(* IEC 61131-3 sources: tgbot_base/CodeSys, 8 files *)

(* ---- GVL_IO.st ---- *)
VAR_GLOBAL
	(* ===================== MODE AND COMMON ===================== *)
	I_ModeManual AT %IX0.0 : BOOL; (* Manual/Automatic selector switch: 1 = Manual, 0 = Automatic *)
	HMI_Auto_Start : BOOL; (* HMI request to enable automatic sequence when in automatic mode *)
	HMI_ResetFaults : BOOL; (* HMI command to reset latched emergency conditions *)

	(* ===================== HMI MANUAL COMMANDS ===================== *)
	HMI_Fan1_Start : BOOL; (* Manual start for Local Fan 1 *)
	HMI_Fan2_Start : BOOL; (* Manual start for Local Fan 2 *)
	HMI_Fan3_Start : BOOL; (* Manual start for Local Fan 3 *)
	HMI_Fan4_Start : BOOL; (* Manual start for Local Fan 4 *)
	HMI_Fan5_Start : BOOL; (* Manual start for Local Fan 5 *)
	HMI_TransportFan_Start : BOOL; (* Manual start for Transport Fan *)
	HMI_Screw_Start : BOOL; (* Manual start for Screw Conveyor *)
	HMI_Vibrator1_Start : BOOL; (* Manual start for Vibrator 1 *)
	HMI_Vibrator2_Start : BOOL; (* Manual start for Vibrator 2 *)
	HMI_Hydraulic_Open : BOOL; (* Manual open command for Hydraulic Hatch *)
	HMI_Hydraulic_Close : BOOL; (* Manual close command for Hydraulic Hatch *)

	(* ===================== PHYSICAL INPUTS (FAULTS, LIMITS) ===================== *)
	(* VFD Faults for Local Fans *)
	I_Fan1_VFD_Fault AT %IX1.0 : BOOL; (* VFD fault for Local Fan 1 *)
	I_Fan2_VFD_Fault AT %IX1.1 : BOOL; (* VFD fault for Local Fan 2 *)
	I_Fan3_VFD_Fault AT %IX1.2 : BOOL; (* VFD fault for Local Fan 3 *)
	I_Fan4_VFD_Fault AT %IX1.3 : BOOL; (* VFD fault for Local Fan 4 *)
	I_Fan5_VFD_Fault AT %IX1.4 : BOOL; (* VFD fault for Local Fan 5 *)

	(* VFD Faults for other mechanisms — keep within byte 1 for example mapping *)
	I_TransportFan_VFD_Fault AT %IX1.5 : BOOL; (* VFD fault for Transport Fan *)
	I_Screw_VFD_Fault AT %IX1.6 : BOOL; (* VFD fault for Screw Conveyor *)
	I_Vibrator1_VFD_Fault AT %IX1.7 : BOOL; (* VFD fault for Vibrator 1 (if applicable) *)
	I_Vibrator2_VFD_Fault AT %IX3.0 : BOOL; (* VFD fault for Vibrator 2 (if applicable); mapped to input byte 3 bit 0 *)

	(* Circuit breaker trips (as per requirement: only vibrators and hydraulic motor) *)
	I_Vibrator1_CB_Trip AT %IX2.0 : BOOL; (* Circuit breaker trip for Vibrator 1 *)
	I_Vibrator2_CB_Trip AT %IX2.1 : BOOL; (* Circuit breaker trip for Vibrator 2 *)
	I_Hydraulic_CB_Trip AT %IX2.2 : BOOL; (* Circuit breaker trip for Hydraulic Power Unit/Motor *)

	(* Hydraulic hatch limit switches *)
	I_Hatch_Open_LS AT %IX2.3 : BOOL; (* Hydraulic Hatch OPEN position limit switch *)
	I_Hatch_Closed_LS AT %IX2.4 : BOOL; (* Hydraulic Hatch CLOSED position limit switch *)

	(* ===================== PHYSICAL OUTPUTS (COMMANDS) ===================== *)
	Q_Fan1_Run AT %QX0.0 : BOOL; (* Run command for Local Fan 1 *)
	Q_Fan2_Run AT %QX0.1 : BOOL; (* Run command for Local Fan 2 *)
	Q_Fan3_Run AT %QX0.2 : BOOL; (* Run command for Local Fan 3 *)
	Q_Fan4_Run AT %QX0.3 : BOOL; (* Run command for Local Fan 4 *)
	Q_Fan5_Run AT %QX0.4 : BOOL; (* Run command for Local Fan 5 *)
	Q_TransportFan_Run AT %QX0.5 : BOOL; (* Run command for Transport Fan *)
	Q_Screw_Run AT %QX0.6 : BOOL; (* Run command for Screw Conveyor *)
	Q_Vibrator1_Run AT %QX1.0 : BOOL; (* Run command for Vibrator 1 *)
	Q_Vibrator2_Run AT %QX1.1 : BOOL; (* Run command for Vibrator 2 *)
	Q_Hydraulic_Open AT %QX1.2 : BOOL; (* Open command for Hydraulic Hatch actuator *)
	Q_Hydraulic_Close AT %QX1.3 : BOOL; (* Close command for Hydraulic Hatch actuator *)

	(* ===================== STATUS / DIAGNOSTICS FOR HMI ===================== *)
	Status_ModeManual : BOOL; (* Current mode: TRUE = Manual, FALSE = Automatic *)
	Status_AutoEnabled : BOOL; (* Auto sequence enable status *)
	Status_EmergencyActive : BOOL; (* Emergency latch active *)

	Status_Fan1_Running : BOOL; (* Status of Local Fan 1 command *)
	Status_Fan2_Running : BOOL; (* Status of Local Fan 2 command *)
	Status_Fan3_Running : BOOL; (* Status of Local Fan 3 command *)
	Status_Fan4_Running : BOOL; (* Status of Local Fan 4 command *)
	Status_Fan5_Running : BOOL; (* Status of Local Fan 5 command *)
	Status_TransportFan_Running : BOOL; (* Status of Transport Fan command *)
	Status_Screw_Running : BOOL; (* Status of Screw Conveyor command *)
	Status_Vibrator1_Running : BOOL; (* Status of Vibrator 1 command *)
	Status_Vibrator2_Running : BOOL; (* Status of Vibrator 2 command *)
	Status_Hydraulic_Busy : BOOL; (* Hydraulic Hatch actuator active (open or close) *)
END_VAR

(* ---- FB_AutoControl.st ---- *)
FUNCTION_BLOCK FB_AutoControl
VAR_INPUT
	AutoMode : BOOL; (* TRUE when selector is in automatic mode *)
	AutoStartRequest : BOOL; (* HMI request to enable automatic sequence *)
	GlobalPermit : BOOL; (* Permit from emergency handling; must be TRUE to run *)
END_VAR
VAR_OUTPUT
	AutoEnabled : BOOL; (* Auto mode active and permitted *)
	Fan1Start : BOOL; (* Auto start command for Local Fan 1 *)
	Fan2Start : BOOL; (* Auto start command for Local Fan 2 *)
	Fan3Start : BOOL; (* Auto start command for Local Fan 3 *)
	Fan4Start : BOOL; (* Auto start command for Local Fan 4 *)
	Fan5Start : BOOL; (* Auto start command for Local Fan 5 *)
	TransportFanStart : BOOL; (* Auto start command for Transport Fan *)
	ScrewStart : BOOL; (* Auto start command for Screw Conveyor *)
	Vibrator1Start : BOOL; (* Auto start command for Vibrator 1 *)
	Vibrator2Start : BOOL; (* Auto start command for Vibrator 2 *)
END_VAR
VAR
	tFan2 : TON;
	tFan3 : TON;
	tFan4 : TON;
	tFan5 : TON;
	tTransport : TON;
	tScrew : TON;
	tVibrators : TON;
	sequenceEnabled : BOOL;
END_VAR

(* Determine if automatic control is enabled *)
sequenceEnabled := AutoMode AND AutoStartRequest AND GlobalPermit;
AutoEnabled := sequenceEnabled;

(* Progressive start delays for fans 2..5 from AutoEnabled *)
tFan2(IN := sequenceEnabled, PT := T#1S);
tFan3(IN := sequenceEnabled, PT := T#2S);
tFan4(IN := sequenceEnabled, PT := T#3S);
tFan5(IN := sequenceEnabled, PT := T#4S);

Fan1Start := sequenceEnabled;
Fan2Start := sequenceEnabled AND tFan2.Q;
Fan3Start := sequenceEnabled AND tFan3.Q;
Fan4Start := sequenceEnabled AND tFan4.Q;
Fan5Start := sequenceEnabled AND tFan5.Q;

(* Transport fan after all local fans are on *)
tTransport(IN := sequenceEnabled AND tFan5.Q, PT := T#1S);
TransportFanStart := sequenceEnabled AND tTransport.Q;

(* Screw after transport fan is running *)
tScrew(IN := sequenceEnabled AND TransportFanStart, PT := T#1S);
ScrewStart := sequenceEnabled AND tScrew.Q;

(* Vibrators after screw is running; both start together *)
tVibrators(IN := sequenceEnabled AND ScrewStart, PT := T#2S);
Vibrator1Start := sequenceEnabled AND tVibrators.Q;
Vibrator2Start := sequenceEnabled AND tVibrators.Q;
END_FUNCTION_BLOCK

(* ---- FB_Emergency.st ---- *)
FUNCTION_BLOCK FB_Emergency
VAR_INPUT
	ModeManual : BOOL; (* Current mode for information if needed *)
	ResetCmd : BOOL; (* HMI reset command *)
	(* VFD faults - individual inputs *)
	Fan1VfdFault : BOOL;
	Fan2VfdFault : BOOL;
	Fan3VfdFault : BOOL;
	Fan4VfdFault : BOOL;
	Fan5VfdFault : BOOL;
	TransportFanVfdFault : BOOL;
	ScrewVfdFault : BOOL;
	Vibrator1VfdFault : BOOL;
	Vibrator2VfdFault : BOOL;
	(* Circuit breaker trips *)
	Vibrator1CBTrip : BOOL;
	Vibrator2CBTrip : BOOL;
	HydraulicCBTrip : BOOL;
END_VAR
VAR_OUTPUT
	EmergencyActive : BOOL; (* Latch TRUE if any emergency condition present *)
	GlobalPermit : BOOL; (* TRUE when no emergency conditions and not latched *)
END_VAR
VAR
	anyFault : BOOL;
	anyTrip : BOOL;
	fanFaultAggregate : BOOL;
END_VAR

(* Aggregate all configured faults *)
fanFaultAggregate := Fan1VfdFault OR Fan2VfdFault OR Fan3VfdFault OR Fan4VfdFault OR Fan5VfdFault;
anyFault := fanFaultAggregate OR TransportFanVfdFault OR ScrewVfdFault OR Vibrator1VfdFault OR Vibrator2VfdFault;
anyTrip := Vibrator1CBTrip OR Vibrator2CBTrip OR HydraulicCBTrip;

(* Latch on any fault or trip; reset only when ResetCmd and all clear *)
IF EmergencyActive THEN
	IF ResetCmd AND NOT anyFault AND NOT anyTrip THEN
		EmergencyActive := FALSE;
	END_IF
ELSE
	IF anyFault OR anyTrip THEN
		EmergencyActive := TRUE;
	END_IF
END_IF;

GlobalPermit := NOT EmergencyActive;
END_FUNCTION_BLOCK

(* ---- FB_Fan.st ---- *)
FUNCTION_BLOCK FB_Fan
VAR_INPUT
	Enable : BOOL; (* Permit from emergency & interlocks *)
	ManualMode : BOOL; (* TRUE = Manual, FALSE = Automatic *)
	ManualStartCmd : BOOL; (* Manual start command from HMI *)
	AutoStartCmd : BOOL; (* Automatic start command from FB_AutoControl *)
	DriveFault : BOOL; (* Frequency drive fault input for this device *)
END_VAR
VAR_OUTPUT
	CmdRun : BOOL; (* Command to the physical output *)
	StatusRunning : BOOL; (* Mirrors CmdRun for HMI/debug *)
	Inhibited : BOOL; (* TRUE if disabled due to fault or no permit *)
END_VAR

(* Select source of command based on mode, apply permits and faults *)
IF Enable AND NOT DriveFault THEN
	IF ManualMode THEN
		CmdRun := ManualStartCmd;
	ELSE
		CmdRun := AutoStartCmd;
	END_IF
ELSE
	CmdRun := FALSE;
END_IF;

StatusRunning := CmdRun;
Inhibited := NOT Enable OR DriveFault;
END_FUNCTION_BLOCK

(* ---- FB_HydraulicHatch.st ---- *)
FUNCTION_BLOCK FB_HydraulicHatch
VAR_INPUT
	Enable : BOOL; (* Permit from emergency & interlocks *)
	ManualMode : BOOL; (* TRUE = Manual, FALSE = Automatic; automatic is not allowed *)
	ManualOpenCmd : BOOL; (* HMI open command *)
	ManualCloseCmd : BOOL; (* HMI close command *)
	LS_Open : BOOL; (* Limit switch: hatch at OPEN position *)
	LS_Closed : BOOL; (* Limit switch: hatch at CLOSED position *)
	CircuitBreakerTrip : BOOL; (* Circuit breaker trip for hydraulic motor *)
END_VAR
VAR_OUTPUT
	CmdOpen : BOOL; (* Command to open the hatch *)
	CmdClose : BOOL; (* Command to close the hatch *)
	Busy : BOOL; (* TRUE when either open or close command is active *)
	InterlockActive : BOOL; (* TRUE if inhibited due to limits, mode, CB trip or no permit *)
END_VAR

VAR
	localPermit : BOOL;
END_VAR

(* Only manual mode is allowed; apply permits and interlocks *)
localPermit := Enable AND ManualMode AND NOT CircuitBreakerTrip;

CmdOpen := FALSE;
CmdClose := FALSE;

IF localPermit THEN
	IF ManualOpenCmd AND NOT LS_Open THEN
		CmdOpen := TRUE;
	ELSIF ManualCloseCmd AND NOT LS_Closed THEN
		CmdClose := TRUE;
	END_IF
END_IF;

Busy := CmdOpen OR CmdClose;
InterlockActive := NOT localPermit OR (ManualOpenCmd AND LS_Open) OR (ManualCloseCmd AND LS_Closed);
END_FUNCTION_BLOCK

(* ---- FB_ScrewConveyor.st ---- *)
FUNCTION_BLOCK FB_ScrewConveyor
VAR_INPUT
	Enable : BOOL; (* Permit from emergency & interlocks *)
	ManualMode : BOOL; (* TRUE = Manual, FALSE = Automatic *)
	ManualStartCmd : BOOL; (* Manual start command from HMI *)
	AutoStartCmd : BOOL; (* Automatic start command from FB_AutoControl *)
	DriveFault : BOOL; (* Frequency drive fault input for the conveyor *)
END_VAR
VAR_OUTPUT
	CmdRun : BOOL; (* Command to the physical output *)
	StatusRunning : BOOL; (* Mirrors CmdRun for HMI/debug *)
	Inhibited : BOOL; (* TRUE if disabled due to fault or no permit *)
END_VAR

IF Enable AND NOT DriveFault THEN
	IF ManualMode THEN
		CmdRun := ManualStartCmd;
	ELSE
		CmdRun := AutoStartCmd;
	END_IF
ELSE
	CmdRun := FALSE;
END_IF;

StatusRunning := CmdRun;
Inhibited := NOT Enable OR DriveFault;
END_FUNCTION_BLOCK

(* ---- FB_Vibrator.st ---- *)
FUNCTION_BLOCK FB_Vibrator
VAR_INPUT
	Enable : BOOL; (* Permit from emergency & interlocks *)
	ManualMode : BOOL; (* TRUE = Manual, FALSE = Automatic *)
	ManualStartCmd : BOOL; (* Manual start command from HMI *)
	AutoStartCmd : BOOL; (* Automatic start command from FB_AutoControl *)
	DriveFault : BOOL; (* VFD fault input if vibrator uses VFD; otherwise tie FALSE *)
	CircuitBreakerTrip : BOOL; (* Circuit breaker trip input (required) *)
END_VAR
VAR_OUTPUT
	CmdRun : BOOL; (* Command to the physical output *)
	StatusRunning : BOOL; (* Mirrors CmdRun for HMI/debug *)
	Inhibited : BOOL; (* TRUE if disabled due to fault or no permit *)
END_VAR

IF Enable AND NOT DriveFault AND NOT CircuitBreakerTrip THEN
	IF ManualMode THEN
		CmdRun := ManualStartCmd;
	ELSE
		CmdRun := AutoStartCmd;
	END_IF
ELSE
	CmdRun := FALSE;
END_IF;

StatusRunning := CmdRun;
Inhibited := NOT Enable OR DriveFault OR CircuitBreakerTrip;
END_FUNCTION_BLOCK

(* ---- PLC_PRG.st ---- *)
PROGRAM PLC_PRG
VAR
	(* Mode *)
	modeManual : BOOL; (* 1=Manual, 0=Automatic from I_ModeManual *)

	(* Emergency FB and adapter variables *)
	emg : FB_Emergency;
	emgFanFault1 : BOOL;
	emgFanFault2 : BOOL;
	emgFanFault3 : BOOL;
	emgFanFault4 : BOOL;
	emgFanFault5 : BOOL;

	(* Auto control FB *)
	autoCtl : FB_AutoControl;

	(* Fans FB instances *)
	fbFan1 : FB_Fan;
	fbFan2 : FB_Fan;
	fbFan3 : FB_Fan;
	fbFan4 : FB_Fan;
	fbFan5 : FB_Fan;

	(* Transport fan FB instance *)
	fbTransportFan : FB_Fan;

	(* Screw conveyor FB instance *)
	fbScrew : FB_ScrewConveyor;

	(* Vibrators FB instances *)
	fbVib1 : FB_Vibrator;
	fbVib2 : FB_Vibrator;

	(* Hydraulic hatch FB instance *)
	fbHatch : FB_HydraulicHatch;

	(* Internal wires for auto commands *)
	aFan1Start : BOOL;
	aFan2Start : BOOL;
	aFan3Start : BOOL;
	aFan4Start : BOOL;
	aFan5Start : BOOL;
	aTransportStart : BOOL;
	aScrewStart : BOOL;
	aVib1Start : BOOL;
	aVib2Start : BOOL;

	(* Global permit *)
	permitGlobal : BOOL;
END_VAR

(* Mode handling *)
modeManual := I_ModeManual;
Status_ModeManual := modeManual;

(* Emergency handling; map faults individually to avoid arrays in PLC_PRG *)
emgFanFault1 := I_Fan1_VFD_Fault;
emgFanFault2 := I_Fan2_VFD_Fault;
emgFanFault3 := I_Fan3_VFD_Fault;
emgFanFault4 := I_Fan4_VFD_Fault;
emgFanFault5 := I_Fan5_VFD_Fault;

emg(ModeManual := modeManual,
	ResetCmd := HMI_ResetFaults,
	Fan1VfdFault := emgFanFault1,
	Fan2VfdFault := emgFanFault2,
	Fan3VfdFault := emgFanFault3,
	Fan4VfdFault := emgFanFault4,
	Fan5VfdFault := emgFanFault5,
	TransportFanVfdFault := I_TransportFan_VFD_Fault,
	ScrewVfdFault := I_Screw_VFD_Fault,
	Vibrator1VfdFault := I_Vibrator1_VFD_Fault,
	Vibrator2VfdFault := I_Vibrator2_VFD_Fault,
	Vibrator1CBTrip := I_Vibrator1_CB_Trip,
	Vibrator2CBTrip := I_Vibrator2_CB_Trip,
	HydraulicCBTrip := I_Hydraulic_CB_Trip);

permitGlobal := emg.GlobalPermit;
Status_EmergencyActive := emg.EmergencyActive;

(* Automatic control *)
autoCtl(AutoMode := NOT modeManual,
	AutoStartRequest := HMI_Auto_Start,
	GlobalPermit := permitGlobal);

Status_AutoEnabled := autoCtl.AutoEnabled;

(* Cache auto commands for readability *)
aFan1Start := autoCtl.Fan1Start;
aFan2Start := autoCtl.Fan2Start;
aFan3Start := autoCtl.Fan3Start;
aFan4Start := autoCtl.Fan4Start;
aFan5Start := autoCtl.Fan5Start;
aTransportStart := autoCtl.TransportFanStart;
aScrewStart := autoCtl.ScrewStart;
aVib1Start := autoCtl.Vibrator1Start;
aVib2Start := autoCtl.Vibrator2Start;

(* Local Fans 1..5 *)
fbFan1(Enable := permitGlobal, ManualMode := modeManual, ManualStartCmd := HMI_Fan1_Start, AutoStartCmd := aFan1Start, DriveFault := I_Fan1_VFD_Fault);
Q_Fan1_Run := fbFan1.CmdRun;
Status_Fan1_Running := fbFan1.StatusRunning;

fbFan2(Enable := permitGlobal, ManualMode := modeManual, ManualStartCmd := HMI_Fan2_Start, AutoStartCmd := aFan2Start, DriveFault := I_Fan2_VFD_Fault);
Q_Fan2_Run := fbFan2.CmdRun;
Status_Fan2_Running := fbFan2.StatusRunning;

fbFan3(Enable := permitGlobal, ManualMode := modeManual, ManualStartCmd := HMI_Fan3_Start, AutoStartCmd := aFan3Start, DriveFault := I_Fan3_VFD_Fault);
Q_Fan3_Run := fbFan3.CmdRun;
Status_Fan3_Running := fbFan3.StatusRunning;

fbFan4(Enable := permitGlobal, ManualMode := modeManual, ManualStartCmd := HMI_Fan4_Start, AutoStartCmd := aFan4Start, DriveFault := I_Fan4_VFD_Fault);
Q_Fan4_Run := fbFan4.CmdRun;
Status_Fan4_Running := fbFan4.StatusRunning;

fbFan5(Enable := permitGlobal, ManualMode := modeManual, ManualStartCmd := HMI_Fan5_Start, AutoStartCmd := aFan5Start, DriveFault := I_Fan5_VFD_Fault);
Q_Fan5_Run := fbFan5.CmdRun;
Status_Fan5_Running := fbFan5.StatusRunning;

(* Transport Fan *)
fbTransportFan(Enable := permitGlobal, ManualMode := modeManual, ManualStartCmd := HMI_TransportFan_Start, AutoStartCmd := aTransportStart, DriveFault := I_TransportFan_VFD_Fault);
Q_TransportFan_Run := fbTransportFan.CmdRun;
Status_TransportFan_Running := fbTransportFan.StatusRunning;

(* Screw Conveyor *)
fbScrew(Enable := permitGlobal, ManualMode := modeManual, ManualStartCmd := HMI_Screw_Start, AutoStartCmd := aScrewStart, DriveFault := I_Screw_VFD_Fault);
Q_Screw_Run := fbScrew.CmdRun;
Status_Screw_Running := fbScrew.StatusRunning;

(* Vibrators *)
fbVib1(Enable := permitGlobal, ManualMode := modeManual, ManualStartCmd := HMI_Vibrator1_Start, AutoStartCmd := aVib1Start, DriveFault := I_Vibrator1_VFD_Fault, CircuitBreakerTrip := I_Vibrator1_CB_Trip);
Q_Vibrator1_Run := fbVib1.CmdRun;
Status_Vibrator1_Running := fbVib1.StatusRunning;

fbVib2(Enable := permitGlobal, ManualMode := modeManual, ManualStartCmd := HMI_Vibrator2_Start, AutoStartCmd := aVib2Start, DriveFault := I_Vibrator2_VFD_Fault, CircuitBreakerTrip := I_Vibrator2_CB_Trip);
Q_Vibrator2_Run := fbVib2.CmdRun;
Status_Vibrator2_Running := fbVib2.StatusRunning;

(* Hydraulic Hatch - manual only with interlocks *)
fbHatch(Enable := permitGlobal, ManualMode := modeManual, ManualOpenCmd := HMI_Hydraulic_Open, ManualCloseCmd := HMI_Hydraulic_Close, LS_Open := I_Hatch_Open_LS, LS_Closed := I_Hatch_Closed_LS, CircuitBreakerTrip := I_Hydraulic_CB_Trip);
Q_Hydraulic_Open := fbHatch.CmdOpen;
Q_Hydraulic_Close := fbHatch.CmdClose;
Status_Hydraulic_Busy := fbHatch.Busy;
END_PROGRAM
